(* IEC 61131-3 sources: Industry-PLC-LLM/data/PLCBEAD_repo/PLCBEAD_PLCEmbed-main/PLC-BEAD/Source/GEB/ESR_MON_X8, 1 file *)

(* ---- ESR_MON_X8.ST ---- *)
TYPE
	oscat_ESR_collect_data      : ARRAY [0..7]    OF BYTE;
END_TYPE

TYPE oscat_ESR_data :
  STRUCT
	typ    : BYTE;
	ADRESS : STRING;
	DS     : UDINT;
	TS     : TIME;
	data   : oscat_ESR_collect_data;
  END_STRUCT;
END_TYPE

TYPE
  oscat_ESR_3                : ARRAY [0..3] OF oscat_ESR_data;
  oscat_ESR_31               : ARRAY [0..31] OF oscat_ESR_data;
END_TYPE

FUNCTION_BLOCK STATUS_TO_ESR_Block

	VAR_INPUT
		STATUS :	BYTE;
		ADRESS :	STRING;
		DT_IN :	UDINT;
		TS :	TIME;
	END_VAR

	VAR_OUTPUT
		STATUS_TO_ESR :	oscat_ESR_data;
	END_VAR

	IF STATUS < BYTE#100 THEN
		STATUS_TO_ESR.typ := BYTE#1;
	ELSIF STATUS < BYTE#200 THEN
		STATUS_TO_ESR.typ := BYTE#2;
	ELSE
		STATUS_TO_ESR.typ := BYTE#3;
	END_IF;
	STATUS_TO_ESR.ADRESS:= ADRESS;
	STATUS_TO_ESR.DS := DT_IN;
	STATUS_TO_ESR.TS := TS;
	STATUS_TO_ESR.data[0] := STATUS;
END_FUNCTION_BLOCK

FUNCTION_BLOCK T_PLC_MS_block

	VAR_OUTPUT
		T_PLC_MS :	UDINT;
	END_VAR

	VAR
		PLC_TICKS_PER_SEC :	INT;
		PLC_SYS_TICK_CNT :	DINT;
	END_VAR

	VAR
		debug :	BOOL;(*Debug-Mode ON / OFF*)
		N :	INT;(*Debug-Faktor*)
		Offset :	UDINT;(*Debug-Offset*)
		temp :	DWORD := DWORD#1;(*Debug-Offset*)
		MODE :	BOOL;(*modus*)
		faktor :	UDINT;(*Systemtakt-Faktor*)
		init :	BOOL;
		v_plc_ticks_per_sec :	UDINT;
		base :	UDINT := UDINT#1000;
	END_VAR

	IF init = FALSE THEN
		v_plc_ticks_per_sec := INT_TO_UDINT(PLC_TICKS_PER_SEC);
		IF v_plc_ticks_per_sec = UDINT#1024 THEN
			faktor := UDINT#1;
			MODE := FALSE;
		ELSIF v_plc_ticks_per_sec > UDINT#0 THEN
			IF v_plc_ticks_per_sec <= base THEN
				faktor := base / v_plc_ticks_per_sec;
				MODE := FALSE;
			ELSE
				faktor := v_plc_ticks_per_sec / base;
				MODE := TRUE;
			END_IF;
		ELSE
			faktor := UDINT#1;
		END_IF;
		init := TRUE;
	END_IF;

	IF MODE THEN
		T_PLC_MS := DINT_TO_UDINT(PLC_SYS_TICK_CNT) / faktor;
	ELSE
		T_PLC_MS := DINT_TO_UDINT(PLC_SYS_TICK_CNT) * faktor;
	END_IF;

	IF debug THEN
		T_PLC_MS := (DWORD_TO_UDINT(SHL(UDINT_TO_DWORD(T_PLC_MS),N) OR SHL(temp,N)) - UDINT#1) + Offset;
	END_IF;

END_FUNCTION_BLOCK

FUNCTION_BLOCK ESR_MON_X8
	VAR_INPUT
		S0 :	BYTE;
		A0 :	STRING;
		S1 :	BYTE;
		A1 :	STRING;
		S2 :	BYTE;
		A2 :	STRING;
		S3 :	BYTE;
		A3 :	STRING;
		S4 :	BYTE;
		A4 :	STRING;
		S5 :	BYTE;
		A5 :	STRING;
		S6 :	BYTE;
		A6 :	STRING;
		S7 :	BYTE;
		A7 :	STRING;
		DT_IN :	UDINT;
		MODE :	BYTE := BYTE#3;
	END_VAR

	VAR_IN_OUT
		ESR_OUT :	oscat_ESR_3;
	END_VAR

	VAR_OUTPUT
		ESR_FLAG :	BOOL;
	END_VAR

	VAR
		X0 :	BYTE;
		X1 :	BYTE;
		X2 :	BYTE;
		X3 :	BYTE;
		X4 :	BYTE;
		X5 :	BYTE;
		X6 :	BYTE;
		X7 :	BYTE;
		TX :	TIME;
		CNT :	INT;
		STATUS_TO_ESR :	STATUS_TO_ESR_Block;
		T_PLC_MS :	T_PLC_MS_block;
	END_VAR

	T_PLC_MS();
	TX:= UDINT_TO_TIME(T_PLC_MS.T_PLC_MS);

	ESR_FLAG := FALSE;
	ESR_OUT[3].typ := BYTE#0;
	ESR_OUT[2].typ := BYTE#0;
	ESR_OUT[1].typ := BYTE#0;
	ESR_OUT[0].typ := BYTE#0;
	CNT := 0;

	IF S0 <> X0 AND ((S0 < BYTE#100) OR (S0 > BYTE#99 AND S0 < BYTE#200 AND MODE >= BYTE#2) OR (S0 > BYTE#199 AND MODE = BYTE#3)) THEN

		STATUS_TO_ESR.STATUS := S0;
		STATUS_TO_ESR.ADRESS := A0;
		STATUS_TO_ESR.DT_IN  := DT_IN;
		STATUS_TO_ESR.TS     := TX;
		STATUS_TO_ESR();
		ESR_OUT[CNT] := STATUS_TO_ESR.STATUS_TO_ESR;

		X0 := S0;
		CNT := CNT + 1;
		ESR_FLAG := TRUE;
	END_IF;
	IF S1 <> X1 AND ((S1 < BYTE#100) OR (S1 > BYTE#99 AND S1 < BYTE#200 AND MODE >= BYTE#2) OR (S1 > BYTE#199 AND MODE = BYTE#3)) THEN

		STATUS_TO_ESR.STATUS := S1;
		STATUS_TO_ESR.ADRESS := A1;
		STATUS_TO_ESR.DT_IN  := DT_IN;
		STATUS_TO_ESR.TS     := TX;
		STATUS_TO_ESR();
		ESR_OUT[CNT] := STATUS_TO_ESR.STATUS_TO_ESR;

		X1 := S1;
		CNT := CNT + 1;
		ESR_FLAG := TRUE;
	END_IF;
	IF S2 <> X2 AND ((S2 < BYTE#100) OR (S2 > BYTE#99 AND S2 < BYTE#200 AND MODE >= BYTE#2) OR (S2 > BYTE#199 AND MODE = BYTE#3)) THEN

		STATUS_TO_ESR.STATUS := S2;
		STATUS_TO_ESR.ADRESS := A2;
		STATUS_TO_ESR.DT_IN  := DT_IN;
		STATUS_TO_ESR.TS     := TX;
		STATUS_TO_ESR();
		ESR_OUT[CNT] := STATUS_TO_ESR.STATUS_TO_ESR;

		X2 := S2;
		CNT := CNT + 1;
		ESR_FLAG := TRUE;
	END_IF;
	IF S3 <> X3 AND ((S3 < BYTE#100) OR (S3 > BYTE#99 AND S3 < BYTE#200 AND MODE >= BYTE#2) OR (S3 > BYTE#199 AND MODE = BYTE#3)) THEN

		STATUS_TO_ESR.STATUS := S3;
		STATUS_TO_ESR.ADRESS := A3;
		STATUS_TO_ESR.DT_IN  := DT_IN;
		STATUS_TO_ESR.TS     := TX;
		STATUS_TO_ESR();
		ESR_OUT[CNT] := STATUS_TO_ESR.STATUS_TO_ESR;

		X3 := S3;
		CNT := CNT + 1;
		ESR_FLAG := TRUE;
	END_IF;
	IF CNT < 4 AND S4 <> X4 AND ((S4 < BYTE#100) OR (S4 > BYTE#99 AND S4 < BYTE#200 AND MODE >= BYTE#2) OR (S4 > BYTE#199 AND MODE = BYTE#3)) THEN

		STATUS_TO_ESR.STATUS := S4;
		STATUS_TO_ESR.ADRESS := A4;
		STATUS_TO_ESR.DT_IN  := DT_IN;
		STATUS_TO_ESR.TS     := TX;
		STATUS_TO_ESR();
		ESR_OUT[CNT] := STATUS_TO_ESR.STATUS_TO_ESR;

		X4 := S4;
		CNT := CNT + 1;
		ESR_FLAG := TRUE;
	END_IF;
	IF CNT < 4 AND S5 <> X5 AND ((S5 < BYTE#100) OR (S5 > BYTE#99 AND S5 < BYTE#200 AND MODE >= BYTE#2) OR (S5 > BYTE#199 AND MODE = BYTE#3)) THEN

		STATUS_TO_ESR.STATUS := S5;
		STATUS_TO_ESR.ADRESS := A5;
		STATUS_TO_ESR.DT_IN  := DT_IN;
		STATUS_TO_ESR.TS     := TX;
		STATUS_TO_ESR();
		ESR_OUT[CNT] := STATUS_TO_ESR.STATUS_TO_ESR;

		X5 := S5;
		CNT := CNT + 1;
		ESR_FLAG := TRUE;
	END_IF;
	IF CNT < 4 AND S6 <> X6 AND ((S6 < BYTE#100) OR (S6 > BYTE#99 AND S6 < BYTE#200 AND MODE >= BYTE#2) OR (S6 > BYTE#199 AND MODE = BYTE#3)) THEN

		STATUS_TO_ESR.STATUS := S6;
		STATUS_TO_ESR.ADRESS := A6;
		STATUS_TO_ESR.DT_IN  := DT_IN;
		STATUS_TO_ESR.TS     := TX;
		STATUS_TO_ESR();
		ESR_OUT[CNT] := STATUS_TO_ESR.STATUS_TO_ESR;

		X6 := S6;
		CNT := CNT + 1;
		ESR_FLAG := TRUE;
	END_IF;
	IF CNT < 4 AND S7 <> X7 AND ((S7 < BYTE#100) OR (S7 > BYTE#99 AND S7 < BYTE#200 AND MODE >= BYTE#2) OR (S7 > BYTE#199 AND MODE = BYTE#3)) THEN

		STATUS_TO_ESR.STATUS := S7;
		STATUS_TO_ESR.ADRESS := A7;
		STATUS_TO_ESR.DT_IN  := DT_IN;
		STATUS_TO_ESR.TS     := TX;
		STATUS_TO_ESR();
		ESR_OUT[CNT] := STATUS_TO_ESR.STATUS_TO_ESR;

		X7 := S7;
		CNT := CNT + 1;
		ESR_FLAG := TRUE;
	END_IF;

END_FUNCTION_BLOCK

PROGRAM program0

	VAR
	S0 :	BYTE;
	A0 :	STRING;
	S1 :	BYTE;
	A1 :	STRING;
	S2 :	BYTE;
	A2 :	STRING;
	S3 :	BYTE;
	A3 :	STRING;
	S4 :	BYTE;
	A4 :	STRING;
	S5 :	BYTE;
	A5 :	STRING;
	S6 :	BYTE;
	A6 :	STRING;
	S7 :	BYTE;
	A7 :	STRING;
	DT_IN :	UDINT;
	MODE :	BYTE;

	ESR_OUT :	oscat_ESR_3;

	ESR_FLAG :	BOOL;

		func_block : ESR_MON_X8;
  	END_VAR
	func_block.S0 := S0;
	func_block.A0 := A0;
	func_block.S1 := S1;
	func_block.A1 := A1;
	func_block.S2 := S2;
	func_block.A2 := A2;
	func_block.S3 := S3;
	func_block.A3 := A3;
	func_block.S4 := S4;
	func_block.A4 := A4;
	func_block.S5 := S5;
	func_block.A5 := A5;
	func_block.S6 := S6;
	func_block.A6 := A6;
	func_block.S7 := S7;
	func_block.A7 := A7;
	func_block.DT_IN := DT_IN;
	func_block.MODE := MODE;
	func_block(ESR_OUT := ESR_OUT);
	ESR_OUT := func_block.ESR_OUT;
	ESR_FLAG := func_block.ESR_FLAG;
END_PROGRAM
